(* IEC 61131-3 sources: stratumak/tests/modcompile-st, 31 files *)

(* ---- actions.st ---- *)
{attribute 'summary' := 'Named pieces of a body, shared with it'}
{attribute 'license' := 'GPL'}

(* An ACTION is a named piece of a POU's body.  It shares every variable of the
   POU and has none of its own, which is what makes it different from a
   FUNCTION_BLOCK: nothing has to be passed in, and nothing has its own state.

   The alternative for splitting a long cyclic body is a function block, which
   changes the state layout and forces every touched variable through an
   interface, or a FUNCTION, which cannot see the POU's variables at all. *)

FUNCTION_BLOCK Counter
  VAR_INPUT
    step  : DINT;
    reset : BOOL;
  END_VAR
  VAR_OUTPUT
    total : DINT;
  END_VAR
  VAR
    overflows : DINT;
  END_VAR

  IF reset THEN
    clear();
  ELSE
    accumulate();
  END_IF;

(* An action of a function block reaches the instance, so its signature is the
   block body's exactly. *)
ACTION clear:
  total := 0;
  overflows := 0;
END_ACTION

ACTION accumulate:
  total := total + step;
  IF total > 1000 THEN
    overflows := overflows + 1;
    clear();
  END_IF;
END_ACTION

END_FUNCTION_BLOCK

{attribute 'doc' := 'Runs the counter and reports on it.'}
PROGRAM actions
  VAR_INPUT
    enable : BOOL;
    amount : DINT := 1;
  END_VAR
  VAR_OUTPUT
    count   : DINT;
    running : BOOL;
    idle    : BOOL;
  END_VAR
  VAR
    c        : Counter;
    selected : DINT;
  END_VAR

  (* An action of an instance, called from outside the block that declares
     it: `motor.stop()`.  It shares that instance's variables and takes no
     arguments -- there is no interface to pass anything through. *)
  c.clear();

  IF enable THEN
    (* An action of a PROGRAM sees the pin snapshot, so it may read and write
       pins exactly as the body does. *)
    advance(selected := amount);
  ELSE
    stop();
  END_IF;

  report();

ACTION advance:
  c(step := selected, reset := FALSE);
  count := c.total;
  running := TRUE;
END_ACTION

ACTION stop:
  c(step := 0, reset := TRUE);
  count := 0;
  running := FALSE;
END_ACTION

(* This one touches no pin at all, only instance state. *)
ACTION report:
  idle := NOT running;
END_ACTION

END_PROGRAM

(* ---- atmap.st ---- *)
{attribute 'summary' := 'Explicit pin mapping with AT'}
{attribute 'license' := 'GPL'}

(* A function block that publishes one of its own values to HAL.  It is not a
   VAR_INPUT, so nothing at a call site writes it -- the direction in the AT
   clause is the whole story, and there is no second writer to conflict with. *)

FUNCTION_BLOCK Axis
  VAR_INPUT
    cmd : LREAL;
  END_VAR
  VAR
    pos AT %Q.position : LREAL;
    err AT %Q.error    : LREAL;
    home AT %I.at_home : BOOL;
  END_VAR

  IF home THEN
    pos := 0.0;
  ELSE
    pos := pos + (cmd - pos) * 0.1;
  END_IF;
  err := cmd - pos;
END_FUNCTION_BLOCK

PROGRAM atmap
  VAR
    (* A plain VAR mapped explicitly, and renamed on the way out. *)
    enable  AT %I         : BOOL;
    running AT %Q.active  : BOOL;
    feed    AT %IO        : LREAL;

    x    : Axis;
    axes : ARRAY[0..2] OF Axis;
    i    : DINT;
  END_VAR

  running := enable;
  x(cmd := feed);
  FOR i := 0 TO 2 DO
    axes[i](cmd := feed);
  END_FOR;
END_PROGRAM

(* ---- bad_extaction.st ---- *)
(* An action has no interface, so a call to one from outside takes no
   arguments.  Inside the declaring POU `Act(v := x)` is shorthand for setting
   one of the POU's own variables first; from outside the same spelling would
   reach past the instance's interface into its state.

   It is also the spelling an IEC ed.3 METHOD call uses, and a syntax whose
   meaning depended on which of the two the name turned out to be would be a
   poor thing to have built. *)

FUNCTION_BLOCK Motor
  VAR_OUTPUT
    speed : DINT;
  END_VAR

  speed := speed;

ACTION stop:
  speed := 0;
END_ACTION

END_FUNCTION_BLOCK

PROGRAM bad_extaction
  VAR_OUTPUT
    q : DINT;
  END_VAR
  VAR
    m : Motor;
  END_VAR

  m.stop(speed := 5);
  q := m.speed;
END_PROGRAM

(* ---- bad_recursive.st ---- *)
{attribute 'summary' := 'A function block that contains itself'}

(* This must be refused.  A block holding an instance of itself is infinitely
   large before it ever runs, and recursion has no place in a real-time body
   anyway: the stack depth cannot be bounded.
   See docs/dev/MODCOMPILE_ST_FRONTEND.md §4. *)

FUNCTION_BLOCK Nested
  VAR_INPUT
    trigger : BOOL;
  END_VAR
  VAR_OUTPUT
    depth : DINT;
  END_VAR
  VAR
    inner : Nested;
  END_VAR

  inner(trigger := trigger);
  depth := inner.depth + 1;
END_FUNCTION_BLOCK

PROGRAM bad_recursive
  VAR_INPUT
    go : BOOL;
  END_VAR
  VAR_OUTPUT
    level : DINT;
  END_VAR
  VAR
    n : Nested;
  END_VAR

  n(trigger := go);
  level := n.depth;
END_PROGRAM

(* ---- bad_thisrec.st ---- *)
(* Until a method could reach a sibling, methods could not recurse at all:
   reaching one needed THIS, and reaching another block's method needed
   containment, which is refused.  Both routes exist now, so the cycle check
   has to see them -- the real-time stack is fixed and there is no useful way
   to bound the depth. *)

FUNCTION_BLOCK Loop
  VAR_OUTPUT
    o : DINT;
  END_VAR

  o := a();

METHOD a : DINT
  a := b();
END_METHOD

METHOD b : DINT
  b := THIS^.a();
END_METHOD

END_FUNCTION_BLOCK

PROGRAM bad_thisrec
  VAR_OUTPUT
    q : DINT;
  END_VAR
  VAR
    l : Loop;
  END_VAR

  l();
  q := l.o;
END_PROGRAM

(* ---- durations.st ---- *)
{attribute 'summary' := 'The TIME type: literals, arithmetic and conversions'}
{attribute 'license' := 'GPL'}

(* A duration is held as int64 nanoseconds -- what get_time() and a task's
   period already are.  It is not a number: it adds to and compares with
   another duration, scales by a count, and divides by another duration to give
   their ratio, and anything else is refused rather than guessed at.

   See docs/dev/MODCOMPILE_ST_STDLIB.md §5. *)

TYPE Config : STRUCT
  (* The shape the production sources actually use: PT is read from a struct
     member far more often than it is written as a literal. *)
  errDelay  : TIME;
  pumpOff   : TIME;
END_STRUCT
END_TYPE

FUNCTION_BLOCK Elapsed
  VAR_INPUT
    run : BOOL;
  END_VAR
  VAR_OUTPUT
    et : TIME;
  END_VAR

  IF run THEN
    (* fperiod is LREAL seconds, so the bridge is named for seconds. *)
    et := et + SECONDS_TO_TIME(fperiod);
  ELSE
    et := T#0s;
  END_IF;
END_FUNCTION_BLOCK

PROGRAM durations
  VAR_INPUT
    run : BOOL;
    (* HAL has no duration type, so a settable one arrives as seconds. *)
    delay_s : LREAL;
  END_VAR
  VAR_OUTPUT
    expired    : BOOL;
    elapsed_ms : DINT;
    remaining  : LREAL;
    fraction   : LREAL;
  END_VAR
  VAR
    cfg : Config;
    e   : Elapsed;

    pt      : TIME := T#500ms;
    warmup  : TIME := T#1m30s;
    fine    : TIME := T#1s500ms250us;
    half    : TIME;
  END_VAR

  cfg.errDelay := SECONDS_TO_TIME(delay_s);
  cfg.pumpOff  := T#2s;

  e(run := run);

  expired    := e.et >= pt;
  elapsed_ms := TIME_TO_DINT(e.et);
  remaining  := TIME_TO_SECONDS(warmup - e.et);
  fraction   := e.et / pt;

  (* Scaling: by a whole count and by a fraction. *)
  half := pt / 2;
  pt   := half * 2;
  warmup := warmup * 1.5;

  IF cfg.errDelay > cfg.pumpOff THEN
    pt := fine;
  END_IF;
END_PROGRAM

(* ---- fbnest.st ---- *)
{attribute 'summary' := 'Nested and arrayed function block instances'}
{attribute 'license' := 'GPL'}

(* A function block instance nests as a struct inside inst_t, so an FB may
   contain another, and an array of instances is unremarkable -- neither
   would be true if instances carried HAL identities of their own. *)

FUNCTION_BLOCK Accumulator
  VAR_INPUT
    add   : LREAL;
    clear : BOOL;
  END_VAR
  VAR_OUTPUT
    total : LREAL;
  END_VAR

  IF clear THEN
    total := 0.0;
  ELSE
    total := total + add;
  END_IF;
END_FUNCTION_BLOCK

FUNCTION_BLOCK Averager
  VAR_INPUT
    sample : LREAL;
    reset  : BOOL;
  END_VAR
  VAR_OUTPUT
    mean : LREAL;
  END_VAR
  VAR
    acc   : Accumulator;
    count : DINT;
  END_VAR

  IF reset THEN
    count := 0;
  ELSE
    count := count + 1;
  END_IF;

  acc(add := sample, clear := reset);

  IF count > 0 THEN
    mean := acc.total / count;
  ELSE
    mean := 0.0;
  END_IF;
END_FUNCTION_BLOCK

PROGRAM fbnest
  VAR_INPUT
    ch    : ARRAY[0..3] OF LREAL;
    reset : BOOL;
  END_VAR
  VAR_OUTPUT
    mean0 : LREAL;
    mean1 : LREAL;
  END_VAR
  VAR
    avg : ARRAY[0..3] OF Averager;
    i   : DINT;
  END_VAR

  FOR i := 0 TO 3 DO
    avg[i](sample := ch[i], reset := reset);
  END_FOR;

  mean0 := avg[0].mean;
  mean1 := avg[1].mean;
END_PROGRAM

(* ---- methods.st ---- *)
{attribute 'summary' := 'Methods on a function block instance'}
{attribute 'license' := 'GPL'}

(* A METHOD is an operation on an instance: it has its own interface and its
   own locals, and it can reach the instance's variables.  That is what makes
   it different from an ACTION, which shares the POU's variables and has no
   interface at all -- and why both can share the `inst.name()` call syntax
   without either having to know about the other.

   See docs/dev/MODCOMPILE_ST_STDLIB.md §7a. *)

FUNCTION_BLOCK Accumulator
  VAR_OUTPUT
    total : DINT;
  END_VAR
  VAR
    calls : DINT;
  END_VAR

  calls := calls + 1;

  (* The block's own body reaching one of its methods, IEC's way round. *)
  IF calls = 1 THEN
    THIS^.clear();
  END_IF;

{attribute 'doc' := 'Add a weighted value and report the new total.'}
METHOD add : DINT
  VAR_INPUT
    n      : DINT;
    weight : DINT;
  END_VAR
  VAR
    (* A method's own local, which does not persist between calls -- that is
       what the block's VAR is for. *)
    scaled : DINT;
  END_VAR

  scaled := n * weight;
  total  := total + scaled;
  add    := total;
END_METHOD

{attribute 'doc' := 'Add one, at the standard weight.'}
METHOD tick : DINT
  (* A sibling method, called with no name for the instance: there is one in
     scope either way, and the generated function already has it. *)
  tick := add(n := 1, weight := 1);
END_METHOD

{attribute 'doc' := 'Start again.'}
METHOD clear
  (* No result type at all: a method that only acts on the instance returns
     nothing, and writing `: VOID` for that would need a type ST does not
     have. *)
  total := 0;
END_METHOD

(* An action beside the methods, sharing the block's variables and taking no
   interface of its own. *)
ACTION note:
  calls := calls + 1;
END_ACTION

END_FUNCTION_BLOCK

PROGRAM methods
  VAR_INPUT
    reset : BOOL;
  END_VAR
  VAR_OUTPUT
    running : DINT;
  END_VAR
  VAR
    acc : Accumulator;
  END_VAR

  acc();

  (* As an expression, for the result... *)
  running := acc.add(n := 5, weight := 2);

  (* ...and as a statement, where there is none to use. *)
  IF reset THEN
    acc.clear();
  END_IF;

  (* The same spelling reaches an action, which is the point of §7a. *)
  acc.note();
END_PROGRAM

(* ---- params.st ---- *)
{attribute 'summary' := 'HAL parameters, at the top level and inside a block'}
{attribute 'license' := 'GPL'}

(* A HAL parameter is a value in shared memory that no signal connects to.
   `AT %MRW` is a tunable HAL sets and the component reads; `AT %MR` is a
   diagnostic the component writes and HAL only reads.  See §3.5. *)

FUNCTION_BLOCK Limiter
  VAR_INPUT
    raw : LREAL;
  END_VAR
  VAR_OUTPUT
    limited : LREAL;
  END_VAR
  VAR
    (* A parameter inside a block becomes one per instance, named by the
       path that reaches it -- exactly as a published pin is. *)
    ceiling AT %MRW        : LREAL := 100.0;
    hits    AT %MR.clamped : DINT;
  END_VAR

  limited := raw;
  IF limited > ceiling THEN
    limited := ceiling;
    hits := hits + 1;
  END_IF;
END_FUNCTION_BLOCK

PROGRAM params
  VAR_INPUT
    cmd : LREAL;
  END_VAR
  VAR_OUTPUT
    out : LREAL;
  END_VAR
  VAR
    {attribute 'doc' := 'Multiplies the command before limiting.'}
    gain    AT %MRW       : LREAL := 1.0;
    {attribute 'doc' := 'Set when the last cycle was scaled down.'}
    scaled  AT %MR.active : BOOL;
    invert  AT %MRW       : BOOL;

    lim : Limiter;
  END_VAR

  lim(raw := cmd * gain);
  out := lim.limited;
  IF invert THEN
    out := -out;
  END_IF;
  scaled := gain < 1.0;
END_PROGRAM

(* ---- period.st ---- *)
{attribute 'summary' := 'fperiod, in each kind of body that may use it'}
{attribute 'license' := 'GPL'}

(* fperiod is the period of the thread this body is running in.  The backend
   reaches it two ways -- from the HAL function's own argument where that is in
   scope, and from the RT task otherwise -- and they are the same number,
   because a HAL function is invoked by its own thread.  See
   docs/dev/MODCOMPILE_ST_STDLIB.md §4. *)

FUNCTION_BLOCK Integrator
  VAR_INPUT
    rate : LREAL;
  END_VAR
  VAR_OUTPUT
    total : LREAL;
  END_VAR

  (* A block body is its own C function and was never handed the argument. *)
  IF rate = 0.0 THEN
    reset();
  ELSE
    total := total + rate * fperiod;
  END_IF;

ACTION reset:
  total := 0.0;
END_ACTION

END_FUNCTION_BLOCK

PROGRAM period
  VAR_INPUT
    enable : BOOL;
    rate   : LREAL;
  END_VAR
  VAR_OUTPUT
    total   : LREAL;
    elapsed : LREAL;
  END_VAR
  VAR
    acc : Integrator;
  END_VAR

  IF enable THEN
    (* An exported body has the argument. *)
    elapsed := elapsed + fperiod;
    acc(rate := rate);
  ELSE
    stop();
  END_IF;
  total := acc.total;

(* An action is its own C function too, even inside a PROGRAM. *)
ACTION stop:
  elapsed := 0.0;
END_ACTION

END_PROGRAM

(* ---- ramplimit.st ---- *)
{attribute 'summary' := 'Rate-limited position follower'}
{attribute 'license' := 'GPL'}
{attribute 'author'  := 'stratuMAK'}

(* The worked example of docs/dev/MODCOMPILE_ST_FRONTEND.md §3.  A function
   block is internal: Ramp has no HAL identity, only ramplimit's own
   VAR_INPUT/VAR_OUTPUT become pins.  Where a sub-component's input should be
   wirable, declare the pin at PROGRAM level and pass it in -- which is what
   `target := target` does here. *)

FUNCTION_BLOCK Ramp
  VAR_INPUT
    target : LREAL;
    rate   : LREAL;
    dt     : LREAL;
  END_VAR
  VAR_OUTPUT
    out    : LREAL;
  END_VAR
  VAR
    step   : LREAL;
  END_VAR

  step := rate * dt;
  IF target > out + step THEN
    out := out + step;
  ELSIF target < out - step THEN
    out := out - step;
  ELSE
    out := target;
  END_IF;
END_FUNCTION_BLOCK

PROGRAM ramplimit
  VAR_INPUT
    {attribute 'doc' := 'Commanded position.'}
    target   : LREAL;
    {attribute 'doc' := 'Maximum rate of change, units per second.'}
    max_rate : LREAL := 10.0;
    enable   : BOOL;
  END_VAR
  VAR_OUTPUT
    out      : LREAL;
  END_VAR
  VAR
    r : Ramp;
  END_VAR

  IF enable THEN
    r(target := target, rate := max_rate, dt := fperiod);
    out := r.out;
  ELSE
    out := target;
  END_IF;
END_PROGRAM

(* ---- strings.st ---- *)
{attribute 'summary' := 'String functions in every kind of body'}
{attribute 'license' := 'GPL'}

FUNCTION_BLOCK Tagger
  VAR_INPUT
    go : BOOL;
  END_VAR
  VAR_OUTPUT
    tag : STRING[32];
  END_VAR
  VAR
    (* A STRING member with an initialiser: a char array, so the block's
       initialiser has to copy it rather than assign it. *)
    base : STRING[8] := 'ax';
  END_VAR

  IF go THEN
    build();
  END_IF

  (* An action and a method each become their own C function, so each needs
     its own buffers -- and a helper either of them calls has to be defined
     in the file whether or not the block's own body calls one. *)
  ACTION build:
    tag := CONCAT(base, '-run');
  END_ACTION

  METHOD suffix : INT
    VAR_INPUT
      extra : STRING[8];
    END_VAR
    tag := CONCAT(base, extra);
    suffix := LEN(tag);
  END_METHOD
END_FUNCTION_BLOCK

FUNCTION shorten : INT
  VAR_INPUT
    s : STRING[32];
  END_VAR
  VAR
    (* A STRING local of a function: declared with its length, and
       initialised at the declaration, which is the one place C takes a
       literal for an array. *)
    cut : STRING[16] := 'none';
  END_VAR
  cut := LEFT(s, 4);
  shorten := LEN(cut);
END_FUNCTION

PROGRAM strings
  VAR_OUTPUT
    n : INT;
  END_VAR
  VAR
    t : Tagger;
    (* A STRING has no HAL representation, so it stays inside the
       component -- which is where a message being assembled belongs. *)
    label : STRING[64];
  END_VAR

  t(go := TRUE);
  n := t.suffix(extra := '!') + shorten(t.tag);
  (* Nested, which is the shape these appear in: each call site gets a
     buffer of its own, so the inner one is not overwritten while the outer
     one is still reading it. *)
  label := CONCAT(CONCAT('tag=', t.tag), '!');
END_PROGRAM

(* ---- timers.st ---- *)
{attribute 'library' := 'timers'}
{attribute 'summary' := 'IEC 61131-3 delay timers'}
{attribute 'license' := 'GPL'}

(* A library: TYPE, FUNCTION and FUNCTION_BLOCK declarations and no PROGRAM,
   marked by the 'library' attribute.  What it declares is generated into the
   consumer's own module -- see docs/dev/MODCOMPILE_ST_STDLIB.md §2 -- so a
   call to one of these blocks is a static C function in the same translation
   unit, checked against this declaration and mapped back here by #line. *)

{attribute 'doc' := 'Delay on: Q follows IN, but only after PT.'}
FUNCTION_BLOCK TON
  VAR_INPUT
    {attribute 'doc' := 'The signal to delay.'}
    IN : BOOL;
    {attribute 'doc' := 'How long IN must stay true before Q follows.'}
    PT : TIME;
  END_VAR
  VAR_OUTPUT
    {attribute 'doc' := 'True once IN has been true for PT.'}
    Q  : BOOL;
    ET : TIME;
  END_VAR

  IF IN THEN
    IF ET < PT THEN
      ET := ET + SECONDS_TO_TIME(fperiod);
    END_IF;
    Q := ET >= PT;
  ELSE
    ET := T#0s;
    Q := FALSE;
  END_IF;
END_FUNCTION_BLOCK

(* Nothing in the tree uses this one.  It must not reach the generated C: a
   block body is a static function and cmods build with -Werror, and a library
   exists precisely to declare more than any one consumer wants. *)
FUNCTION_BLOCK TOF
  VAR_INPUT
    IN : BOOL;
    PT : TIME;
  END_VAR
  VAR_OUTPUT
    Q : BOOL;
  END_VAR

  Q := IN OR PT > T#0s;
END_FUNCTION_BLOCK

(* ---- and2.st ---- *)
{attribute 'summary' := 'Two-input AND gate'}
{attribute 'license' := 'GPL'}
{attribute 'author'  := 'stratuMAK'}

(* The smallest useful component: two inputs, one output, no state.
   The .comp equivalent is src/hal/components/and2.comp. *)

PROGRAM and2
  VAR_INPUT
    {attribute 'doc' := 'First input.'}
    in0 : BOOL;
    {attribute 'doc' := 'Second input.'}
    in1 : BOOL;
  END_VAR
  VAR_OUTPUT
    {attribute 'doc' := 'TRUE when both inputs are TRUE.'}
    out : BOOL;
  END_VAR

  out := in0 AND in1;
END_PROGRAM

(* ---- arrays.st ---- *)
{attribute 'summary' := 'Select and average from an array pin'}
{attribute 'license' := 'GPL'}

(* Array pins map one dimension only, since a HAL pin name carries one
   index: channel.0 .. channel.7.  Multi-dimensional arrays are fine as
   internal state.  The non-zero lower bound on `window` is deliberate --
   every index site has to subtract it. *)

PROGRAM arrays
  VAR_INPUT
    channel  : ARRAY[0..7] OF LREAL;
    selected : DINT := 0;
  END_VAR
  VAR_OUTPUT
    value   : LREAL;
    average : LREAL;
  END_VAR
  VAR
    window : ARRAY[1..4] OF LREAL;
    grid   : ARRAY[0..1, 0..2] OF LREAL;
    total  : LREAL;
    i, j   : DINT;
  END_VAR

  value := channel[selected];

  total := 0.0;
  FOR i := 0 TO 7 DO
    total := total + channel[i];
  END_FOR;
  average := total / 8.0;

  FOR i := 1 TO 4 DO
    window[i] := average;
  END_FOR;

  FOR i := 0 TO 1 DO
    FOR j := 0 TO 2 DO
      grid[i, j] := average;
    END_FOR;
  END_FOR;
END_PROGRAM

(* ---- bad_action.st ---- *)
(* An action calling itself is recursion by another name: the stack depth
   cannot be bounded, so the real-time rules refuse it exactly as they refuse a
   recursive FUNCTION. *)

PROGRAM bad_action
  VAR_OUTPUT
    out : DINT;
  END_VAR

  spin();

ACTION spin:
  out := out + 1;
  spin();
END_ACTION

END_PROGRAM

(* ---- bad_address.st ---- *)
{attribute 'summary' := 'An IEC physical address in an AT clause'}

(* This must be refused.  %QX0.0 is a physical address -- memory area, size
   code, offset -- and stratuMAK has no address space to locate a variable in,
   because HAL signals are the addressing scheme.  Saying so beats an
   "unknown direction" that leaves the author guessing.
   See docs/dev/MODCOMPILE_ST_FRONTEND.md §3.1. *)

PROGRAM bad_address
  VAR
    lamp AT %QX0.0 : BOOL;
  END_VAR

  lamp := TRUE;
END_PROGRAM

(* ---- bad_cname.st ---- *)
(* Every variable, pin, parameter and struct field reaches the generated C as
   a bare identifier, so one named for a C keyword would produce code the C
   compiler rejects -- an error against generated source nobody keeps, which is
   the whole thing this frontend exists to prevent. *)

PROGRAM bad_cname
  VAR_OUTPUT
    q : DINT;
  END_VAR
  VAR
    int : DINT;
  END_VAR

  int := 1;
  q := int;
END_PROGRAM

(* ---- bad_index.st ---- *)
{attribute 'summary' := 'A constant subscript outside the declared bounds'}

(* An index the compiler can see is a mistake, not something to clamp: this
   must be refused at compile time.  A subscript it cannot see is clamped at
   run time instead -- see arrays.st. *)

PROGRAM bad_index
  VAR_INPUT
    value : DINT;
  END_VAR
  VAR_OUTPUT
    out : DINT;
  END_VAR
  VAR
    slots : ARRAY[1..4] OF DINT;
  END_VAR

  slots[5] := value;
  out := slots[1];
END_PROGRAM

(* ---- bad_library.st ---- *)
(* A library that is not there.  The message lists every directory searched,
   because that is the question being asked. *)

USING nosuchlibrary;

PROGRAM bad_library
  VAR_OUTPUT
    q : BOOL;
  END_VAR

  q := TRUE;
END_PROGRAM

(* ---- bad_param.st ---- *)
(* An rw parameter is HAL's to set and the component's to read, which is the
   same division an input pin has -- so writing one is refused for the same
   reason.  A component that wants to clamp a tunable reads it and keeps the
   clamped value in a VAR. *)

PROGRAM bad_param
  VAR_OUTPUT
    out : LREAL;
  END_VAR
  VAR
    gain AT %MRW : LREAL := 1.0;
  END_VAR

  IF gain > 10.0 THEN
    gain := 10.0;
  END_IF;
  out := gain;
END_PROGRAM

(* ---- bad_period.st ---- *)
(* A stateless FUNCTION that depended on the rate of whatever thread called it
   would not be stateless, so fperiod is not available in one.  IEC's own
   analog blocks take CYCLE as an explicit input for the same reason. *)

FUNCTION scale : LREAL
  VAR_INPUT
    v : LREAL;
  END_VAR

  scale := v * fperiod;
END_FUNCTION

PROGRAM bad_period
  VAR_OUTPUT
    out : LREAL;
  END_VAR

  out := scale(1.0);
END_PROGRAM

(* ---- bad_pinlen.st ---- *)
(* HAL stores a name in STMAK_HAL_NAME_LEN characters, and truncates anything
   longer.  Two pins differing only past that become one pin on the machine and
   nothing says so, which is why this is refused here instead.

   An array pin is measured at its widest element: what has to fit is
   bad_pinlen.<name>.99, not bad_pinlen.<name>. *)

PROGRAM bad_pinlen
  VAR_OUTPUT
    zzzzzzzzzzzzzzzzzzzzzzzzzzzzzzzzzzzzzzzzzzzzzzzzzzzzzzzzzzzzzzzzzzzzzzzzzzzzzzzzzzzzzzzzzzzzzzzzzzzzzzzzzzzzzzzzzzzzzzzzzzzz : ARRAY [0..99] OF DINT;
  END_VAR

  zzzzzzzzzzzzzzzzzzzzzzzzzzzzzzzzzzzzzzzzzzzzzzzzzzzzzzzzzzzzzzzzzzzzzzzzzzzzzzzzzzzzzzzzzzzzzzzzzzzzzzzzzzzzzzzzzzzzzzzzzzzz[0] := 1;
END_PROGRAM

(* ---- bad_shared_name.st ---- *)
{attribute 'summary' := 'Two programs claiming one name'}

(* This must be refused.  The PROGRAMs of one file share a single instance and
   a single HAL component, so two of them cannot both declare a pin called
   `ready` -- the second registration would collide at load time. *)

PROGRAM read
  VAR_INPUT
    raw : DINT;
  END_VAR
  VAR_OUTPUT
    ready : BOOL;
  END_VAR

  ready := raw > 0;
END_PROGRAM

PROGRAM write
  VAR_INPUT
    gain : DINT;
  END_VAR
  VAR_OUTPUT
    ready : BOOL;
  END_VAR

  ready := gain > 0;
END_PROGRAM

(* ---- bad_time.st ---- *)
(* A duration is not a number.  Adding one to it would be adding one what?
   The combinations that have an unambiguous meaning are accepted and the rest
   are refused by name, rather than guessed at. *)

PROGRAM bad_time
  VAR_OUTPUT
    out : BOOL;
  END_VAR
  VAR
    pt : TIME := T#500ms;
  END_VAR

  pt := pt + 1;
  out := pt > T#0s;
END_PROGRAM

(* ---- bad_unbounded.st ---- *)
{attribute 'summary' := 'A loop with no bound the compiler can see'}

(* This must be refused: a WHILE in a HAL function body has to carry an
   explicit max_iterations cap, because it runs in the real-time thread.
   See docs/dev/MODCOMPILE_ST_FRONTEND.md §4. *)

PROGRAM bad_unbounded
  VAR_INPUT
    limit : DINT;
  END_VAR
  VAR_OUTPUT
    done : BOOL;
  END_VAR
  VAR
    n : DINT;
  END_VAR

  WHILE n < limit DO
    n := n + 1;
  END_WHILE;

  done := n >= limit;
END_PROGRAM

(* ---- documented.st ---- *)
{attribute 'summary'     := 'Every documentation field, exercised'}
{attribute 'description' := 'A component that exists to prove its man page is as complete as one generated from a .comp: description, function docs, per-pin docs, notes, examples, author, licence and see-also.'}
{attribute 'license'     := 'GPL'}
{attribute 'author'      := 'stratuMAK'}
{attribute 'see_also'    := '\fBscale\fR(9), \fBand2\fR(9).'}
{attribute 'notes'       := 'The two functions may run in different threads; only \fBupdate\fR needs a floating-point one.'}
{attribute 'examples'    := 'loadrt documented$Naddf documented.sample servo-thread$Naddf documented.update servo-thread'}

(* Metadata before the first declaration describes the component.  A pragma
   heading a PROGRAM documents that program's HAL function, and one inside a
   VAR section documents the pin it precedes. *)

VAR_GLOBAL
  latest : DINT;
END_VAR

{attribute 'doc' := 'Latches the raw input when strobed. Uses no floating point.'}
PROGRAM sample
  VAR_INPUT
    {attribute 'doc' := 'Value to latch.'}
    raw : DINT;
    {attribute 'doc' := 'Rising level latches \fBraw\fR.'}
    strobe : BOOL;
  END_VAR
  VAR_OUTPUT
    {attribute 'doc' := 'TRUE once a value has been latched.'}
    valid : BOOL;
  END_VAR

  IF strobe THEN
    latest := raw;
    valid := TRUE;
  END_IF;
END_PROGRAM

{attribute 'doc' := 'Scales the latched value. Requires a floating-point thread.'}
PROGRAM update
  VAR_INPUT
    {attribute 'doc' := 'Multiplier applied to the latched value.'}
    gain : LREAL := 1.0;
  END_VAR
  VAR_OUTPUT
    {attribute 'doc' := 'The latched value times \fBgain\fR.'}
    scaled : LREAL;
  END_VAR

  scaled := latest * gain;
END_PROGRAM

(* ---- loops.st ---- *)
{attribute 'summary' := 'Bounded iteration'}
{attribute 'license' := 'GPL'}

(* Every loop in a HAL function body carries a bound the compiler can see.
   FOR is bounded by construction.  WHILE and REPEAT are not, so each needs
   an explicit max_iterations cap -- without one, sema rejects the statement.
   See docs/dev/MODCOMPILE_ST_FRONTEND.md §4. *)

PROGRAM loops
  VAR_INPUT
    target    : LREAL;
    tolerance : LREAL := 0.001;
  END_VAR
  VAR_OUTPUT
    estimate   : LREAL;
    iterations : DINT;
  END_VAR
  VAR
    guess : LREAL;
    i     : DINT;
  END_VAR

  guess := target / 2.0;
  iterations := 0;

  (* Newton-Raphson for a square root: iterative settling is a real pattern,
     and a bounded WHILE says so more honestly than a FOR with a break. *)
  {attribute 'max_iterations' := '50'}
  WHILE guess * guess - target > tolerance DO
    guess := (guess + target / guess) / 2.0;
    iterations := iterations + 1;
  END_WHILE;

  {attribute 'max_iterations' := '10'}
  REPEAT
    iterations := iterations + 1;
  UNTIL iterations > 5
  END_REPEAT;

  FOR i := 0 TO 9 DO
    IF i > 4 THEN
      EXIT;
    END_IF;
    iterations := iterations + 1;
  END_FOR;

  estimate := guess;
END_PROGRAM

(* ---- statemachine.st ---- *)
{attribute 'summary' := 'Three-state sequencer with a fault path'}
{attribute 'license' := 'GPL'}

(* An enumeration used as a state variable, with CASE arms labelled by
   constant name rather than by number.  Resolving those names is exactly
   what the standalone prototype could not do. *)

TYPE
  State : (IDLE, RUNNING, FAULTED);
END_TYPE

PROGRAM statemachine
  VAR_INPUT
    start   : BOOL;
    stop    : BOOL;
    fault   : BOOL;
    reset   : BOOL;
  END_VAR
  VAR_OUTPUT
    is_running : BOOL;
    alarm   : BOOL;
  END_VAR
  VAR
    state : State := IDLE;
  END_VAR

  IF fault THEN
    state := FAULTED;
  END_IF;

  CASE state OF
    IDLE:
      IF start AND NOT stop THEN
        state := RUNNING;
      END_IF;
    RUNNING:
      IF stop THEN
        state := IDLE;
      END_IF;
    FAULTED:
      IF reset AND NOT fault THEN
        state := IDLE;
      END_IF;
  ELSE
    state := FAULTED;
  END_CASE;

  is_running := state = RUNNING;
  alarm   := state = FAULTED;
END_PROGRAM

(* ---- twoprograms.st ---- *)
{attribute 'summary' := 'Two thread functions sharing state'}
{attribute 'license' := 'GPL'}

(* One PROGRAM per exported HAL function.  These become twoprograms.read and
   twoprograms.write, addf-able to different threads, with VAR_GLOBAL the
   state they share.  Each PROGRAM carries its own pins.

   `read` touches no floating point, so it should export with fp = 0. *)

VAR_GLOBAL
  latched : DINT;
  ready   : BOOL;
END_VAR

PROGRAM read
  VAR_INPUT
    raw    : DINT;
    strobe : BOOL;
  END_VAR
  VAR_OUTPUT
    accepted : BOOL;
  END_VAR

  IF strobe THEN
    latched := raw;
    ready := TRUE;
  END_IF;
  accepted := ready;
END_PROGRAM

PROGRAM write
  VAR_INPUT
    gain : LREAL := 1.0;
  END_VAR
  VAR_OUTPUT
    scaled : LREAL;
    valid  : BOOL;
  END_VAR

  IF ready THEN
    scaled := latched * gain;
    valid  := TRUE;
  ELSE
    scaled := 0.0;
    valid  := FALSE;
  END_IF;
END_PROGRAM

(* ---- uselib.st ---- *)
{attribute 'summary' := 'Uses the timers library'}
{attribute 'license' := 'GPL'}

USING timers;

PROGRAM uselib
  VAR_INPUT
    start : BOOL;
  END_VAR
  VAR_OUTPUT
    running : BOOL;
    elapsed : LREAL;
  END_VAR
  VAR
    delay : TON;
  END_VAR

  delay(IN := start, PT := T#500ms);
  running := delay.Q;
  elapsed := TIME_TO_SECONDS(delay.ET);
END_PROGRAM
